(* IEC 61131-3 sources: PLC-Static-Analysis/modules/plc-rules/src/test/resources/PLCA-L019, 2 files *)

(* ---- compliant.st ---- *)
PROGRAM P_L019ok
VAR
    n : INT;
    m : INT;
    r : REAL;
    b : BOOL;
    c : BOOL;
    q : BOOL;
END_VAR
IF n > 10 THEN
    q := TRUE;
END_IF
IF n > 10 THEN
    q := TRUE;
ELSE
    b := FALSE;
END_IF
IF n > 10 THEN
    q := TRUE;
ELSE
    q := TRUE;
END_IF
q := n > 10;
END_PROGRAM

(* ---- noncompliant.st ---- *)
PROGRAM P_L019
VAR
    n : INT;
    m : INT;
    r : REAL;
    b : BOOL;
    c : BOOL;
    q : BOOL;
END_VAR
IF n > 10 THEN // PLCA-L019
    q := TRUE;
ELSE
    q := FALSE;
END_IF
IF b AND c THEN // PLCA-L019
    q := FALSE;
ELSE
    q := TRUE;
END_IF
END_PROGRAM
